Staubli VAL3: onSave.pgx

program onSave()
  local bool l_bResult
  local num l_i
begin
  actdata:aActItem[nSelList].sComment=aEditItem.sComment
  for l_i = 0 to size(aEditItem.aActItem)-1
    actdata:aActItem[nSelList].aActItem[l_i].sIOtype=aEditItem.aActItem[l_i].sIOtype
    actdata:aActItem[nSelList].aActItem[l_i].sValue=aEditItem.aActItem[l_i].sValue
    actdata:aActItem[nSelList].aActItem[l_i].bActive=(aEditItem.aActItem[l_i].bActive==true)
    toNum(sSelIO[l_i],actdata:aActItem[nSelList].aActItem[l_i].nIOindex,l_bResult)
    if !l_bResult
      actdata:aActItem[nSelList].aActItem[l_i].nIOindex=-1
    endIf
    actdata:aActItem[nSelList].aActItem[l_i].nPulseValue=aEditItem.aActItem[l_i].nPulseValue
  endFor
  bOnsave=true
  actdata:libSave()
  delay(0.1)
end
